// TIA Portal V20 export
// export: Created 2026-10-19T18:02:05.6879248Z, ExportSetting WithDefaults, DisplayName Totally Integrated Automation Portal, DisplayVersion V20 Update 6, DisplayName TIA Portal Openness, DisplayVersion V20 Update 6, DisplayName TIA Portal Version Control Interface, DisplayVersion V20 Update 6, DisplayName SINAMICS Startdrive Advanced, DisplayVersion V20 SP1, DisplayName SINAMICS Startdrive G130, G150, S120, S150, SINAMICS MV, G220, S200, S210, DisplayVersion V20 SP1, DisplayName SINAMICS Startdrive G110M, G120, G120C, G120D, G120P, G115D, DisplayVersion V20 SP1, DisplayName STEP 7 Professional, DisplayVersion V20 Update 6, DisplayName STEP 7 Safety, DisplayVersion V20 Update 2, DisplayName WinCC Basic/Comfort/Advanced, DisplayVersion V20 Update 6, DisplayName WinCC Unified, DisplayVersion V20 Update 6
FUNCTION_BLOCK "Main_Safety_RTG1"   // FB1, F_FBD
{ S7_Optimized_Access := 'TRUE' }
VERSION : 0.1
// stored: AutoNumber false, IsIECCheckEnabled false, UDAEnableTagReadback false
   VAR
      SAFETY_OK_VTD : Bool;
      SAFETY_OK_CAROUSEL : Bool;
      MAIN_PANEL_OK : Bool;
      REMOTE_PANEL_OK : Bool;
      "E-STOP_INBOUND_OK" : Bool;
      PICK_STATION_OK : Bool;
      data_Safe : DInt;
      "HMI_E-STOP" : Bool;
   END_VAR
BEGIN

REGION Network 1: SAFETY OK VTD
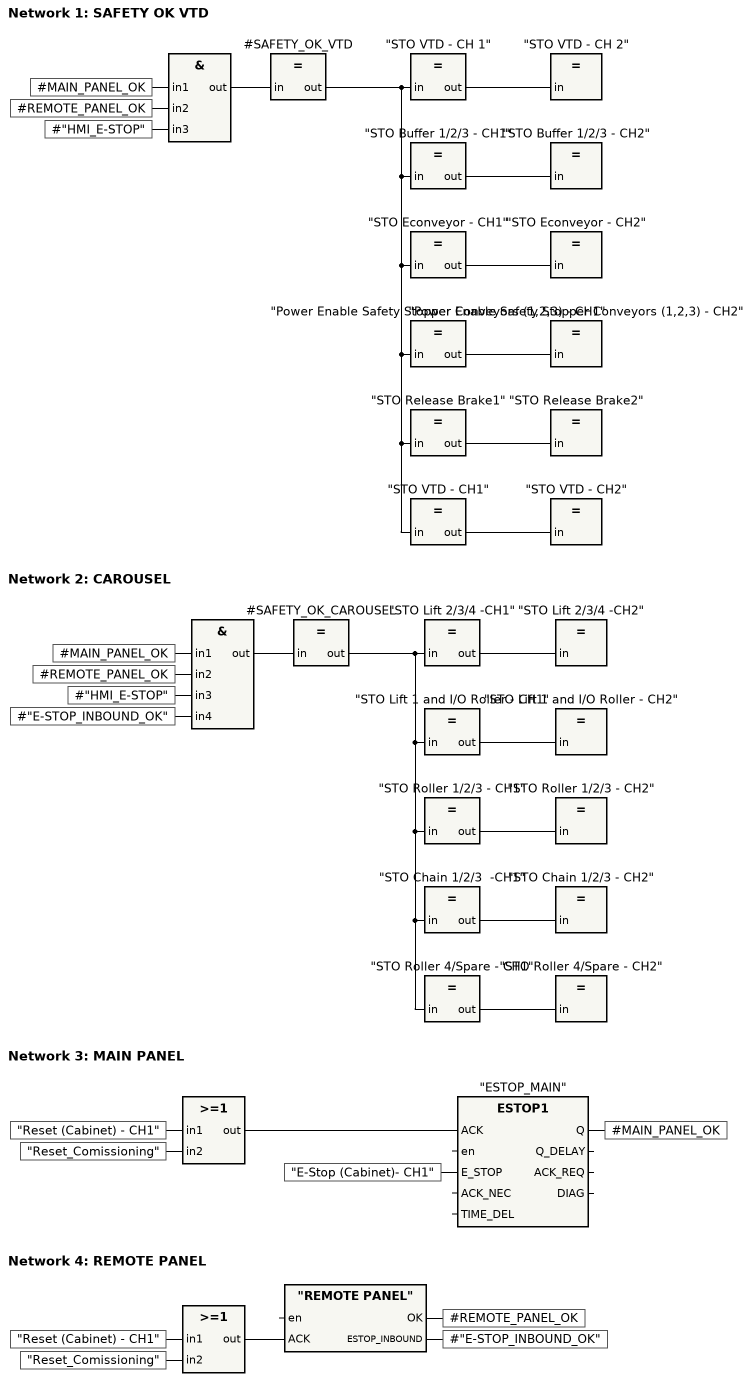
   #SAFETY_OK_VTD := #MAIN_PANEL_OK AND #REMOTE_PANEL_OK AND #"HMI_E-STOP";
   "STO VTD - CH 1" := #SAFETY_OK_VTD;
   "STO VTD - CH 2" := #SAFETY_OK_VTD;
   "STO Buffer 1/2/3 - CH1" := #SAFETY_OK_VTD;
   "STO Buffer 1/2/3 - CH2" := #SAFETY_OK_VTD;
   "STO Econveyor - CH1" := #SAFETY_OK_VTD;
   "STO Econveyor - CH2" := #SAFETY_OK_VTD;
   "Power Enable Safety Stopper Conveyors (1,2,3) - CH1" := #SAFETY_OK_VTD;
   "Power Enable Safety Stopper Conveyors (1,2,3) - CH2" := #SAFETY_OK_VTD;
   "STO Release Brake1" := #SAFETY_OK_VTD;
   "STO Release Brake2" := #SAFETY_OK_VTD;
   "STO VTD - CH1" := #SAFETY_OK_VTD;
   "STO VTD - CH2" := #SAFETY_OK_VTD;
END_REGION

REGION Network 2: CAROUSEL
   #SAFETY_OK_CAROUSEL := #MAIN_PANEL_OK AND #REMOTE_PANEL_OK AND #"HMI_E-STOP" AND #"E-STOP_INBOUND_OK";
   "STO Lift 2/3/4 -CH1" := #SAFETY_OK_CAROUSEL;
   "STO Lift 2/3/4 -CH2" := #SAFETY_OK_CAROUSEL;
   "STO Lift 1 and I/O Roller - CH1" := #SAFETY_OK_CAROUSEL;
   "STO Lift 1 and I/O Roller - CH2" := #SAFETY_OK_CAROUSEL;
   "STO Roller 1/2/3 - CH1" := #SAFETY_OK_CAROUSEL;
   "STO Roller 1/2/3 - CH2" := #SAFETY_OK_CAROUSEL;
   "STO Chain 1/2/3  -CH1" := #SAFETY_OK_CAROUSEL;
   "STO Chain 1/2/3 - CH2" := #SAFETY_OK_CAROUSEL;
   "STO Roller 4/Spare - CH1" := #SAFETY_OK_CAROUSEL;
   "STO Roller 4/Spare - CH2" := #SAFETY_OK_CAROUSEL;
END_REGION

REGION Network 3: MAIN PANEL
   "ESTOP_MAIN"(ACK := "Reset (Cabinet) - CH1" OR "Reset_Comissioning",   // ESTOP1
                E_STOP := "E-Stop (Cabinet)- CH1",
                Q => #MAIN_PANEL_OK);
END_REGION

REGION Network 4: REMOTE PANEL
   "REMOTE PANEL"(ACK := "Reset (Cabinet) - CH1" OR "Reset_Comissioning",
                  OK => #REMOTE_PANEL_OK,
                  ESTOP_INBOUND => #"E-STOP_INBOUND_OK");
END_REGION

REGION Network 5: 1=Acknowledgment for reintegration required
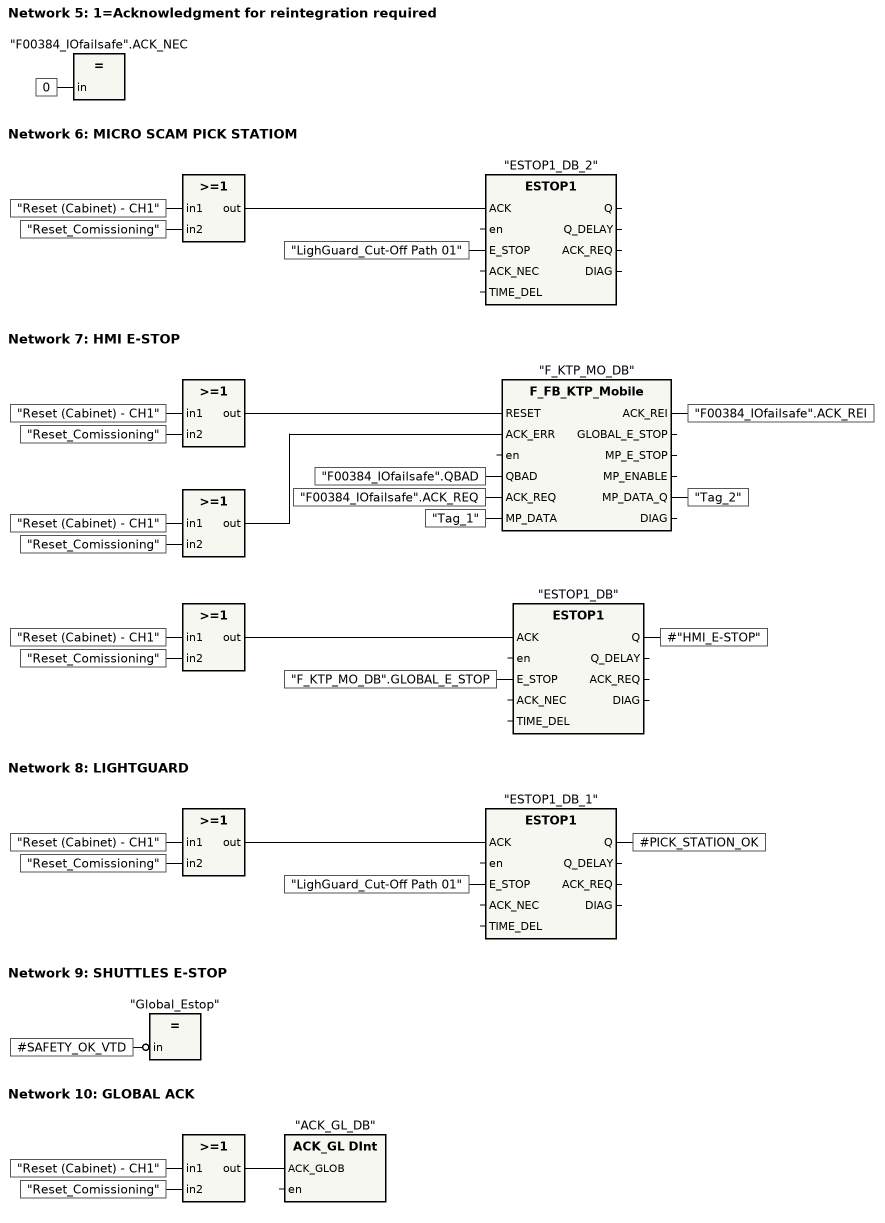
   "F00384_IOfailsafe".ACK_NEC := 0;
END_REGION

REGION Network 6: MICRO SCAM PICK STATIOM
   "ESTOP1_DB_2"(ACK := "Reset (Cabinet) - CH1" OR "Reset_Comissioning", E_STOP := "LighGuard_Cut-Off Path 01");   // ESTOP1
END_REGION

REGION Network 7: HMI E-STOP
   "F_KTP_MO_DB"(RESET := "Reset (Cabinet) - CH1" OR "Reset_Comissioning",   // F_FB_KTP_Mobile
                 ACK_ERR := "Reset (Cabinet) - CH1" OR "Reset_Comissioning",
                 QBAD := "F00384_IOfailsafe".QBAD,
                 ACK_REQ := "F00384_IOfailsafe".ACK_REQ,
                 MP_DATA := "Tag_1",
                 ACK_REI => "F00384_IOfailsafe".ACK_REI,
                 MP_DATA_Q => "Tag_2");
   "ESTOP1_DB"(ACK := "Reset (Cabinet) - CH1" OR "Reset_Comissioning",   // ESTOP1
               E_STOP := "F_KTP_MO_DB".GLOBAL_E_STOP,
               Q => #"HMI_E-STOP");
END_REGION

REGION Network 8: LIGHTGUARD
   "ESTOP1_DB_1"(ACK := "Reset (Cabinet) - CH1" OR "Reset_Comissioning",   // ESTOP1
                 E_STOP := "LighGuard_Cut-Off Path 01",
                 Q => #PICK_STATION_OK);
END_REGION

REGION Network 9: SHUTTLES E-STOP
   "Global_Estop" := NOT #SAFETY_OK_VTD;
END_REGION

REGION Network 10: GLOBAL ACK
   "ACK_GL_DB"(ACK_GLOB := "Reset (Cabinet) - CH1" OR "Reset_Comissioning");   // ACK_GL
END_REGION
END_FUNCTION_BLOCK
